(* IEC 61131-3 sources: codesys-to-s7/tests/corpus/C2S7-PROF-REF/pos, 1 file *)

(* ---- input.st ---- *)
FUNCTION_BLOCK FB_Case
VAR
    r : REFERENCE TO INT;
    a : INT;
END_VAR
r REF= a;
END_FUNCTION_BLOCK
